(* IEC 61131-3 sources: plc-vscode/tests/st/all/trust-platform/manual-tests/root-a/libs/Core, 1 file *)

(* ---- Lib.st ---- *)
NAMESPACE Vendor.Core
FUNCTION CoreFn : DINT
VAR_INPUT X : DINT; END_VAR
CoreFn := X;
END_FUNCTION
END_NAMESPACE
